FUNCTION_BLOCK ServiceTest (* Service interface with request and confirmation *)
  (* Standard: 61499-1; Description: Copyright (c) 2026 Martin Erich Jobst This program and the accompanying materials are made available under the terms of the Eclipse Public License 2.0 which is available at https://www.eclipse.org/legal/epl-2.0/ SPDX-License-Identifier: EPL-2.0 *)
  (* Version 1.0, 2026-10-23, Martin Jobst *)
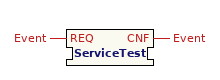
  EVENT_INPUT
    REQ; (* Request *)
  END_EVENT
  EVENT_OUTPUT
    CNF; (* Confirmation *)
  END_EVENT
  SERVICE PLUG/SOCKET (* Request-confirmation service *)
    SEQUENCE request_confirm {SET_ATTRIBUTE(StartState, REQ)} {SET_ATTRIBUTE(ServiceSequenceType, ALWAYS)}
      SOCKET.REQ() -> PLUG.REQ();
      PLUG.CNF() -> SOCKET.CNF();
    END_SEQUENCE
  END_SERVICE
END_FUNCTION_BLOCK
